KUKA KRL data list: MAIN_1.dat

&ACCESS RVP
&REL 1
&COMMENT Generated by RoboDK
&PARAM TEMPLATE = C:\KRC\Roboter\Template\vorgabe
&PARAM EDITMASK = *
DEFDAT  MAIN_1

EXT BAS (BAS_COMMAND :IN,REAL :IN )
EXT REMOTE_PROG_CALL_171()
EXT PICK_PART_111()
EXT PLACE_PART_112()
EXT EVENT_PROG_START_101()
EXT EVENT_PATH_APPROACH_102()
EXT EVENT_PATH_START_103()
EXT EVENT_PATH_FINISH_105()
EXT EVENT_PATH_RETRACT_106()
EXT EVENT_PROG_FINISH_107()
EXT PROG1_withaverylongnameandspecialcharacters()

DECL E6AXIS XP1={A1 -0.00000,A2 0.00000,A3 0.00000,A4 0.00000,A5 0.00000,A6 -0.00000}
DECL FDAT FP1={TOOL_NO 1,BASE_NO 1,IPO_FRAME #BASE,POINT2[] " ",TQ_STATE FALSE}
DECL PDAT PPDAT1={VEL 100.000,ACC 100.000,APO_DIST 1.000,APO_MODE #CPTP}
DECL E6AXIS XP2={A1 0.00000,A2 3.21124,A3 -15.42370,A4 0.00000,A5 12.21250,A6 -0.00000}
DECL FDAT FP2={TOOL_NO 1,BASE_NO 1,IPO_FRAME #BASE,POINT2[] " ",TQ_STATE FALSE}
DECL PDAT PPDAT2={VEL 100.000,ACC 100.000,APO_DIST 1.000,APO_MODE #CPTP}
DECL E6POS XP3={X 1015.000,Y 0.000,Z 1272.000,A 0.000,B 90.000,C 0.000}
DECL FDAT FP3={TOOL_NO 1,BASE_NO 1,IPO_FRAME #BASE,POINT2[] " ",TQ_STATE FALSE}
DECL LDAT LCPDAT3={VEL 1.00000,ACC 100.000,APO_DIST 1.000,APO_FAC 50.0000,ORI_TYP #VAR,CIRC_TYP #BASE,JERK_FAC 50.0000}
DECL E6AXIS XP4={A1 -29.33220,A2 46.67700,A3 -0.02452,A4 26.54560,A5 25.39570,A6 -51.63400}
DECL FDAT FP4={TOOL_NO 1,BASE_NO 1,IPO_FRAME #BASE,POINT2[] " ",TQ_STATE FALSE}
DECL PDAT PPDAT4={VEL 100.000,ACC 100.000,APO_DIST 10.000,APO_MODE #CPTP}
DECL E6POS XP5={X 187.786,Y 125.499,Z 139.112,A -179.997,B 0.180,C 179.996}
DECL FDAT FP5={TOOL_NO 1,BASE_NO 1,IPO_FRAME #BASE,POINT2[] " ",TQ_STATE FALSE}
DECL LDAT LCPDAT5={VEL 0.10000,ACC 100.000,APO_DIST 1.000,APO_FAC 50.0000,ORI_TYP #VAR,CIRC_TYP #BASE,JERK_FAC 50.0000}
DECL E6POS XP6={X 187.272,Y 447.522,Z 305.347,A 179.999,B 0.185,C -179.998}
DECL FDAT FP6={TOOL_NO 1,BASE_NO 1,IPO_FRAME #BASE,POINT2[] " ",TQ_STATE FALSE}
DECL LDAT LCPDAT6={VEL 0.30000,ACC 100.000,APO_DIST 10.000,APO_FAC 50.0000,ORI_TYP #VAR,CIRC_TYP #BASE,JERK_FAC 50.0000}
DECL E6POS XP7={X 187.851,Y 447.517,Z 126.235,A 179.999,B 0.185,C -179.998}
DECL FDAT FP7={TOOL_NO 1,BASE_NO 1,IPO_FRAME #BASE,POINT2[] " ",TQ_STATE FALSE}
DECL LDAT LCPDAT7={VEL 0.10000,ACC 100.000,APO_DIST 1.000,APO_FAC 50.0000,ORI_TYP #VAR,CIRC_TYP #BASE,JERK_FAC 50.0000}
DECL E6POS XP8={X 187.272,Y 447.522,Z 305.347,A 179.999,B 0.185,C -179.998}
DECL FDAT FP8={TOOL_NO 1,BASE_NO 1,IPO_FRAME #BASE,POINT2[] " ",TQ_STATE FALSE}
DECL LDAT LCPDAT8={VEL 0.10000,ACC 100.000,APO_DIST 10.000,APO_FAC 50.0000,ORI_TYP #VAR,CIRC_TYP #BASE,JERK_FAC 50.0000}
DECL E6AXIS XP9={A1 52.18600,A2 45.67580,A3 6.92000,A4 66.73420,A5 19.93230,A6 -92.73000}
DECL FDAT FP9={TOOL_NO 1,BASE_NO 1,IPO_FRAME #BASE,POINT2[] " ",TQ_STATE FALSE}
DECL PDAT PPDAT9={VEL 100.000,ACC 100.000,APO_DIST 25.000,APO_MODE #CPTP}
DECL E6POS XP10={X 430.047,Y 43.774,Z 231.503,A -134.549,B 11.181,C 178.913}
DECL E6POS XP11={X 109.688,Y -153.222,Z 161.073,A -134.549,B 11.181,C 178.913}
DECL FDAT FP11={TOOL_NO 1,BASE_NO 1,IPO_FRAME #BASE,POINT2[] " ",TQ_STATE FALSE}
DECL LDAT LCPDAT11={VEL 0.10000,ACC 100.000,APO_DIST 25.000,APO_FAC 50.0000,ORI_TYP #VAR,CIRC_TYP #BASE,JERK_FAC 50.0000}
DECL E6POS XP12={X 312.208,Y 292.214,Z 255.156,A -134.549,B 11.181,C 178.913}
DECL FDAT FP12={TOOL_NO 1,BASE_NO 1,IPO_FRAME #BASE,POINT2[] " ",TQ_STATE FALSE}
DECL LDAT LCPDAT12={VEL 0.10000,ACC 100.000,APO_DIST 1.000,APO_FAC 50.0000,ORI_TYP #VAR,CIRC_TYP #BASE,JERK_FAC 50.0000}
DECL E6AXIS XP13={A1 -0.00000,A2 0.00000,A3 0.00000,A4 0.00000,A5 0.00000,A6 -0.00000}
DECL FDAT FP13={TOOL_NO 1,BASE_NO 1,IPO_FRAME #BASE,POINT2[] " ",TQ_STATE FALSE}
DECL PDAT PPDAT13={VEL 100.000,ACC 100.000,APO_DIST 1.000,APO_MODE #CPTP}
DECL E6AXIS XP14={A1 88.67600,A2 29.60160,A3 -6.42883,A4 -1.98422,A5 49.47920,A6 4.54769}
DECL FDAT FP14={TOOL_NO 1,BASE_NO 1,IPO_FRAME #BASE,POINT2[] " ",TQ_STATE FALSE}
DECL PDAT PPDAT14={VEL 100.000,ACC 100.000,APO_DIST 1.000,APO_MODE #CPTP}
DECL E6POS XP15={X 19.898,Y 174.307,Z 19.008,A -94.928,B -5.426,C -179.533}
DECL FDAT FP15={TOOL_NO 1,BASE_NO 1,IPO_FRAME #BASE,POINT2[] " ",TQ_STATE FALSE}
DECL LDAT LCPDAT15={VEL 0.10000,ACC 100.000,APO_DIST 1.000,APO_FAC 50.0000,ORI_TYP #VAR,CIRC_TYP #BASE,JERK_FAC 50.0000}
DECL E6POS XP16={X 378.402,Y 174.416,Z 18.997,A -94.928,B -5.426,C -179.533}
DECL FDAT FP16={TOOL_NO 1,BASE_NO 1,IPO_FRAME #BASE,POINT2[] " ",TQ_STATE FALSE}
DECL LDAT LCPDAT16={VEL 0.10000,ACC 100.000,APO_DIST 1.000,APO_FAC 50.0000,ORI_TYP #VAR,CIRC_TYP #BASE,JERK_FAC 50.0000}
DECL E6POS XP17={X 380.996,Y 112.363,Z 34.882,A -95.294,B -18.136,C -178.348}
DECL FDAT FP17={TOOL_NO 1,BASE_NO 1,IPO_FRAME #BASE,POINT2[] " ",TQ_STATE FALSE}
DECL LDAT LCPDAT17={VEL 0.10000,ACC 100.000,APO_DIST 1.000,APO_FAC 50.0000,ORI_TYP #VAR,CIRC_TYP #BASE,JERK_FAC 50.0000}
DECL E6POS XP18={X 16.551,Y 114.359,Z 34.226,A -95.294,B -18.136,C -178.348}
DECL FDAT FP18={TOOL_NO 1,BASE_NO 1,IPO_FRAME #BASE,POINT2[] " ",TQ_STATE FALSE}
DECL LDAT LCPDAT18={VEL 0.10000,ACC 100.000,APO_DIST 1.000,APO_FAC 50.0000,ORI_TYP #VAR,CIRC_TYP #BASE,JERK_FAC 50.0000}
DECL E6POS XP19={X 26.434,Y 54.524,Z 46.072,A -95.461,B 4.348,C 179.585}
DECL FDAT FP19={TOOL_NO 1,BASE_NO 1,IPO_FRAME #BASE,POINT2[] " ",TQ_STATE FALSE}
DECL LDAT LCPDAT19={VEL 0.10000,ACC 100.000,APO_DIST 1.000,APO_FAC 50.0000,ORI_TYP #VAR,CIRC_TYP #BASE,JERK_FAC 50.0000}
DECL E6POS XP20={X 385.448,Y 48.050,Z 45.137,A -95.590,B 11.181,C 178.913}
DECL FDAT FP20={TOOL_NO 1,BASE_NO 1,IPO_FRAME #BASE,POINT2[] " ",TQ_STATE FALSE}
DECL LDAT LCPDAT20={VEL 0.10000,ACC 100.000,APO_DIST 1.000,APO_FAC 50.0000,ORI_TYP #VAR,CIRC_TYP #BASE,JERK_FAC 50.0000}
DECL E6POS XP21={X 385.448,Y -1.625,Z 295.251,A -95.590,B 11.181,C 178.913}
DECL FDAT FP21={TOOL_NO 1,BASE_NO 1,IPO_FRAME #BASE,POINT2[] " ",TQ_STATE FALSE}
DECL LDAT LCPDAT21={VEL 0.10000,ACC 100.000,APO_DIST 1.000,APO_FAC 50.0000,ORI_TYP #VAR,CIRC_TYP #BASE,JERK_FAC 50.0000}
DECL E6AXIS XP22={A1 -0.00000,A2 0.00000,A3 0.00000,A4 0.00000,A5 0.00000,A6 -0.00000}
DECL FDAT FP22={TOOL_NO 1,BASE_NO 1,IPO_FRAME #BASE,POINT2[] " ",TQ_STATE FALSE}
DECL PDAT PPDAT22={VEL 100.000,ACC 100.000,APO_DIST 1.000,APO_MODE #CPTP}
DECL E6AXIS XP23={A1 -68.09030,A2 24.20190,A3 26.78550,A4 38.21340,A5 36.20170,A6 -98.79640}
DECL FDAT FP23={TOOL_NO 1,BASE_NO 1,IPO_FRAME #BASE,POINT2[] " ",TQ_STATE FALSE}
DECL PDAT PPDAT23={VEL 100.000,ACC 100.000,APO_DIST 1.000,APO_MODE #CPTP}
DECL E6POS XP24={X -49.895,Y 253.259,Z 319.999,A -90.000,B 0.353,C -179.975}
DECL FDAT FP24={TOOL_NO 1,BASE_NO 1,IPO_FRAME #BASE,POINT2[] " ",TQ_STATE FALSE}
DECL LDAT LCPDAT24={VEL 1.00000,ACC 100.000,APO_DIST 1.000,APO_FAC 50.0000,ORI_TYP #VAR,CIRC_TYP #BASE,JERK_FAC 50.0000}
DECL E6POS XP25={X 0.000,Y 250.000,Z 270.000,A -90.000,B 0.353,C -179.975}
DECL FDAT FP25={TOOL_NO 1,BASE_NO 1,IPO_FRAME #BASE,POINT2[] " ",TQ_STATE FALSE}
DECL LDAT LCPDAT25={VEL 1.00000,ACC 100.000,APO_DIST 1.000,APO_FAC 50.0000,ORI_TYP #VAR,CIRC_TYP #BASE,JERK_FAC 50.0000}
DECL E6POS XP26={X 35.579,Y 247.455,Z 270.000,A -90.000,B 0.345,C -179.925}
DECL FDAT FP26={TOOL_NO 1,BASE_NO 1,IPO_FRAME #BASE,POINT2[] " ",TQ_STATE FALSE}
DECL LDAT LCPDAT26={VEL 0.05000,ACC 100.000,APO_DIST 1.000,APO_FAC 50.0000,ORI_TYP #VAR,CIRC_TYP #BASE,JERK_FAC 50.0000}
DECL E6POS XP27={X 70.433,Y 239.873,Z 270.000,A -89.999,B 0.331,C -179.876}
DECL FDAT FP27={TOOL_NO 1,BASE_NO 1,IPO_FRAME #BASE,POINT2[] " ",TQ_STATE FALSE}
DECL LDAT LCPDAT27={VEL 0.05000,ACC 100.000,APO_DIST 1.000,APO_FAC 50.0000,ORI_TYP #VAR,CIRC_TYP #BASE,JERK_FAC 50.0000}
DECL E6POS XP28={X 103.854,Y 227.408,Z 270.000,A -89.999,B 0.310,C -179.831}
DECL FDAT FP28={TOOL_NO 1,BASE_NO 1,IPO_FRAME #BASE,POINT2[] " ",TQ_STATE FALSE}
DECL LDAT LCPDAT28={VEL 0.05000,ACC 100.000,APO_DIST 1.000,APO_FAC 50.0000,ORI_TYP #VAR,CIRC_TYP #BASE,JERK_FAC 50.0000}
DECL E6POS XP29={X 135.160,Y 210.313,Z 270.000,A -89.999,B 0.283,C -179.788}
DECL FDAT FP29={TOOL_NO 1,BASE_NO 1,IPO_FRAME #BASE,POINT2[] " ",TQ_STATE FALSE}
DECL LDAT LCPDAT29={VEL 0.05000,ACC 100.000,APO_DIST 1.000,APO_FAC 50.0000,ORI_TYP #VAR,CIRC_TYP #BASE,JERK_FAC 50.0000}
DECL E6POS XP30={X 163.715,Y 188.937,Z 270.000,A -89.999,B 0.250,C -179.750}
DECL FDAT FP30={TOOL_NO 1,BASE_NO 1,IPO_FRAME #BASE,POINT2[] " ",TQ_STATE FALSE}
DECL LDAT LCPDAT30={VEL 0.05000,ACC 100.000,APO_DIST 1.000,APO_FAC 50.0000,ORI_TYP #VAR,CIRC_TYP #BASE,JERK_FAC 50.0000}
DECL E6POS XP31={X 188.937,Y 163.715,Z 270.000,A -89.999,B 0.212,C -179.717}
DECL FDAT FP31={TOOL_NO 1,BASE_NO 1,IPO_FRAME #BASE,POINT2[] " ",TQ_STATE FALSE}
DECL LDAT LCPDAT31={VEL 0.05000,ACC 100.000,APO_DIST 1.000,APO_FAC 50.0000,ORI_TYP #VAR,CIRC_TYP #BASE,JERK_FAC 50.0000}
DECL E6POS XP32={X 210.313,Y 135.160,Z 270.000,A -89.999,B 0.170,C -179.689}
DECL FDAT FP32={TOOL_NO 1,BASE_NO 1,IPO_FRAME #BASE,POINT2[] " ",TQ_STATE FALSE}
DECL LDAT LCPDAT32={VEL 0.05000,ACC 100.000,APO_DIST 1.000,APO_FAC 50.0000,ORI_TYP #VAR,CIRC_TYP #BASE,JERK_FAC 50.0000}
DECL E6POS XP33={X 227.408,Y 103.854,Z 270.000,A -89.999,B 0.124,C -179.668}
DECL FDAT FP33={TOOL_NO 1,BASE_NO 1,IPO_FRAME #BASE,POINT2[] " ",TQ_STATE FALSE}
DECL LDAT LCPDAT33={VEL 0.05000,ACC 100.000,APO_DIST 1.000,APO_FAC 50.0000,ORI_TYP #VAR,CIRC_TYP #BASE,JERK_FAC 50.0000}
DECL E6POS XP34={X 239.873,Y 70.433,Z 270.000,A -90.000,B 0.075,C -179.654}
DECL FDAT FP34={TOOL_NO 1,BASE_NO 1,IPO_FRAME #BASE,POINT2[] " ",TQ_STATE FALSE}
DECL LDAT LCPDAT34={VEL 0.05000,ACC 100.000,APO_DIST 1.000,APO_FAC 50.0000,ORI_TYP #VAR,CIRC_TYP #BASE,JERK_FAC 50.0000}
DECL E6POS XP35={X 247.455,Y 35.579,Z 270.000,A -90.000,B 0.025,C -179.647}
DECL FDAT FP35={TOOL_NO 1,BASE_NO 1,IPO_FRAME #BASE,POINT2[] " ",TQ_STATE FALSE}
DECL LDAT LCPDAT35={VEL 0.05000,ACC 100.000,APO_DIST 1.000,APO_FAC 50.0000,ORI_TYP #VAR,CIRC_TYP #BASE,JERK_FAC 50.0000}
DECL E6POS XP36={X 250.000,Y 0.000,Z 270.000,A -90.000,B -0.025,C -179.647}
DECL FDAT FP36={TOOL_NO 1,BASE_NO 1,IPO_FRAME #BASE,POINT2[] " ",TQ_STATE FALSE}
DECL LDAT LCPDAT36={VEL 0.05000,ACC 100.000,APO_DIST 1.000,APO_FAC 50.0000,ORI_TYP #VAR,CIRC_TYP #BASE,JERK_FAC 50.0000}
DECL E6POS XP37={X 247.455,Y -35.579,Z 270.000,A -90.000,B -0.075,C -179.654}
DECL FDAT FP37={TOOL_NO 1,BASE_NO 1,IPO_FRAME #BASE,POINT2[] " ",TQ_STATE FALSE}
DECL LDAT LCPDAT37={VEL 0.05000,ACC 100.000,APO_DIST 1.000,APO_FAC 50.0000,ORI_TYP #VAR,CIRC_TYP #BASE,JERK_FAC 50.0000}
DECL E6POS XP38={X 239.873,Y -70.433,Z 270.000,A -90.001,B -0.124,C -179.668}
DECL FDAT FP38={TOOL_NO 1,BASE_NO 1,IPO_FRAME #BASE,POINT2[] " ",TQ_STATE FALSE}
DECL LDAT LCPDAT38={VEL 0.05000,ACC 100.000,APO_DIST 1.000,APO_FAC 50.0000,ORI_TYP #VAR,CIRC_TYP #BASE,JERK_FAC 50.0000}
DECL E6POS XP39={X 227.408,Y -103.854,Z 270.000,A -90.001,B -0.170,C -179.689}
DECL FDAT FP39={TOOL_NO 1,BASE_NO 1,IPO_FRAME #BASE,POINT2[] " ",TQ_STATE FALSE}
DECL LDAT LCPDAT39={VEL 0.05000,ACC 100.000,APO_DIST 1.000,APO_FAC 50.0000,ORI_TYP #VAR,CIRC_TYP #BASE,JERK_FAC 50.0000}
DECL E6POS XP40={X 210.313,Y -135.160,Z 270.000,A -90.001,B -0.212,C -179.717}
DECL FDAT FP40={TOOL_NO 1,BASE_NO 1,IPO_FRAME #BASE,POINT2[] " ",TQ_STATE FALSE}
DECL LDAT LCPDAT40={VEL 0.05000,ACC 100.000,APO_DIST 1.000,APO_FAC 50.0000,ORI_TYP #VAR,CIRC_TYP #BASE,JERK_FAC 50.0000}
DECL E6POS XP41={X 188.937,Y -163.715,Z 270.000,A -90.001,B -0.250,C -179.750}
DECL FDAT FP41={TOOL_NO 1,BASE_NO 1,IPO_FRAME #BASE,POINT2[] " ",TQ_STATE FALSE}
DECL LDAT LCPDAT41={VEL 0.05000,ACC 100.000,APO_DIST 1.000,APO_FAC 50.0000,ORI_TYP #VAR,CIRC_TYP #BASE,JERK_FAC 50.0000}
DECL E6POS XP42={X 163.715,Y -188.937,Z 270.000,A -90.001,B -0.283,C -179.788}
DECL FDAT FP42={TOOL_NO 1,BASE_NO 1,IPO_FRAME #BASE,POINT2[] " ",TQ_STATE FALSE}
DECL LDAT LCPDAT42={VEL 0.05000,ACC 100.000,APO_DIST 1.000,APO_FAC 50.0000,ORI_TYP #VAR,CIRC_TYP #BASE,JERK_FAC 50.0000}
DECL E6POS XP43={X 135.160,Y -210.313,Z 270.000,A -90.001,B -0.311,C -179.830}
DECL FDAT FP43={TOOL_NO 1,BASE_NO 1,IPO_FRAME #BASE,POINT2[] " ",TQ_STATE FALSE}
DECL LDAT LCPDAT43={VEL 0.05000,ACC 100.000,APO_DIST 1.000,APO_FAC 50.0000,ORI_TYP #VAR,CIRC_TYP #BASE,JERK_FAC 50.0000}
DECL E6POS XP44={X 103.854,Y -227.408,Z 270.000,A -90.001,B -0.332,C -179.876}
DECL FDAT FP44={TOOL_NO 1,BASE_NO 1,IPO_FRAME #BASE,POINT2[] " ",TQ_STATE FALSE}
DECL LDAT LCPDAT44={VEL 0.05000,ACC 100.000,APO_DIST 1.000,APO_FAC 50.0000,ORI_TYP #VAR,CIRC_TYP #BASE,JERK_FAC 50.0000}
DECL E6POS XP45={X 70.433,Y -239.873,Z 270.000,A -90.000,B -0.346,C -179.925}
DECL FDAT FP45={TOOL_NO 1,BASE_NO 1,IPO_FRAME #BASE,POINT2[] " ",TQ_STATE FALSE}
DECL LDAT LCPDAT45={VEL 0.05000,ACC 100.000,APO_DIST 1.000,APO_FAC 50.0000,ORI_TYP #VAR,CIRC_TYP #BASE,JERK_FAC 50.0000}
DECL E6POS XP46={X 35.579,Y -247.455,Z 270.000,A -90.000,B -0.353,C -179.975}
DECL FDAT FP46={TOOL_NO 1,BASE_NO 1,IPO_FRAME #BASE,POINT2[] " ",TQ_STATE FALSE}
DECL LDAT LCPDAT46={VEL 0.05000,ACC 100.000,APO_DIST 1.000,APO_FAC 50.0000,ORI_TYP #VAR,CIRC_TYP #BASE,JERK_FAC 50.0000}
DECL E6POS XP47={X 0.000,Y -250.000,Z 270.000,A -90.000,B -0.353,C -179.975}
DECL FDAT FP47={TOOL_NO 1,BASE_NO 1,IPO_FRAME #BASE,POINT2[] " ",TQ_STATE FALSE}
DECL LDAT LCPDAT47={VEL 0.05000,ACC 100.000,APO_DIST 1.000,APO_FAC 50.0000,ORI_TYP #VAR,CIRC_TYP #BASE,JERK_FAC 50.0000}
DECL E6POS XP48={X 0.000,Y -250.000,Z 270.000,A -90.000,B -0.353,C 179.975}
DECL FDAT FP48={TOOL_NO 1,BASE_NO 1,IPO_FRAME #BASE,POINT2[] " ",TQ_STATE FALSE}
DECL LDAT LCPDAT48={VEL 0.05000,ACC 100.000,APO_DIST 1.000,APO_FAC 50.0000,ORI_TYP #VAR,CIRC_TYP #BASE,JERK_FAC 50.0000}
DECL E6POS XP49={X -35.579,Y -247.455,Z 270.000,A -90.000,B -0.346,C 179.925}
DECL FDAT FP49={TOOL_NO 1,BASE_NO 1,IPO_FRAME #BASE,POINT2[] " ",TQ_STATE FALSE}
DECL LDAT LCPDAT49={VEL 0.05000,ACC 100.000,APO_DIST 1.000,APO_FAC 50.0000,ORI_TYP #VAR,CIRC_TYP #BASE,JERK_FAC 50.0000}
DECL E6POS XP50={X -70.433,Y -239.873,Z 270.000,A -89.999,B -0.331,C 179.876}
DECL FDAT FP50={TOOL_NO 1,BASE_NO 1,IPO_FRAME #BASE,POINT2[] " ",TQ_STATE FALSE}
DECL LDAT LCPDAT50={VEL 0.05000,ACC 100.000,APO_DIST 1.000,APO_FAC 50.0000,ORI_TYP #VAR,CIRC_TYP #BASE,JERK_FAC 50.0000}
DECL E6POS XP51={X -103.854,Y -227.408,Z 270.000,A -89.999,B -0.310,C 179.831}
DECL FDAT FP51={TOOL_NO 1,BASE_NO 1,IPO_FRAME #BASE,POINT2[] " ",TQ_STATE FALSE}
DECL LDAT LCPDAT51={VEL 0.05000,ACC 100.000,APO_DIST 1.000,APO_FAC 50.0000,ORI_TYP #VAR,CIRC_TYP #BASE,JERK_FAC 50.0000}
DECL E6POS XP52={X -135.160,Y -210.313,Z 270.000,A -89.999,B -0.283,C 179.788}
DECL FDAT FP52={TOOL_NO 1,BASE_NO 1,IPO_FRAME #BASE,POINT2[] " ",TQ_STATE FALSE}
DECL LDAT LCPDAT52={VEL 0.05000,ACC 100.000,APO_DIST 1.000,APO_FAC 50.0000,ORI_TYP #VAR,CIRC_TYP #BASE,JERK_FAC 50.0000}
DECL E6POS XP53={X -163.715,Y -188.937,Z 270.000,A -89.999,B -0.250,C 179.750}
DECL FDAT FP53={TOOL_NO 1,BASE_NO 1,IPO_FRAME #BASE,POINT2[] " ",TQ_STATE FALSE}
DECL LDAT LCPDAT53={VEL 0.05000,ACC 100.000,APO_DIST 1.000,APO_FAC 50.0000,ORI_TYP #VAR,CIRC_TYP #BASE,JERK_FAC 50.0000}
DECL E6POS XP54={X -188.937,Y -163.715,Z 270.000,A -89.999,B -0.212,C 179.717}
DECL FDAT FP54={TOOL_NO 1,BASE_NO 1,IPO_FRAME #BASE,POINT2[] " ",TQ_STATE FALSE}
DECL LDAT LCPDAT54={VEL 0.05000,ACC 100.000,APO_DIST 1.000,APO_FAC 50.0000,ORI_TYP #VAR,CIRC_TYP #BASE,JERK_FAC 50.0000}
DECL E6POS XP55={X -210.313,Y -135.160,Z 270.000,A -89.999,B -0.169,C 179.690}
DECL FDAT FP55={TOOL_NO 1,BASE_NO 1,IPO_FRAME #BASE,POINT2[] " ",TQ_STATE FALSE}
DECL LDAT LCPDAT55={VEL 0.05000,ACC 100.000,APO_DIST 1.000,APO_FAC 50.0000,ORI_TYP #VAR,CIRC_TYP #BASE,JERK_FAC 50.0000}
DECL E6POS XP56={X -227.408,Y -103.854,Z 270.000,A -89.999,B -0.123,C 179.669}
DECL FDAT FP56={TOOL_NO 1,BASE_NO 1,IPO_FRAME #BASE,POINT2[] " ",TQ_STATE FALSE}
DECL LDAT LCPDAT56={VEL 0.05000,ACC 100.000,APO_DIST 1.000,APO_FAC 50.0000,ORI_TYP #VAR,CIRC_TYP #BASE,JERK_FAC 50.0000}
DECL E6POS XP57={X -239.873,Y -70.433,Z 270.000,A -90.000,B -0.075,C 179.654}
DECL FDAT FP57={TOOL_NO 1,BASE_NO 1,IPO_FRAME #BASE,POINT2[] " ",TQ_STATE FALSE}
DECL LDAT LCPDAT57={VEL 0.05000,ACC 100.000,APO_DIST 1.000,APO_FAC 50.0000,ORI_TYP #VAR,CIRC_TYP #BASE,JERK_FAC 50.0000}
DECL E6POS XP58={X -247.455,Y -35.579,Z 270.000,A -90.000,B -0.025,C 179.647}
DECL FDAT FP58={TOOL_NO 1,BASE_NO 1,IPO_FRAME #BASE,POINT2[] " ",TQ_STATE FALSE}
DECL LDAT LCPDAT58={VEL 0.05000,ACC 100.000,APO_DIST 1.000,APO_FAC 50.0000,ORI_TYP #VAR,CIRC_TYP #BASE,JERK_FAC 50.0000}
DECL E6POS XP59={X -250.000,Y 0.000,Z 270.000,A -90.000,B 0.025,C 179.647}
DECL FDAT FP59={TOOL_NO 1,BASE_NO 1,IPO_FRAME #BASE,POINT2[] " ",TQ_STATE FALSE}
DECL LDAT LCPDAT59={VEL 0.05000,ACC 100.000,APO_DIST 1.000,APO_FAC 50.0000,ORI_TYP #VAR,CIRC_TYP #BASE,JERK_FAC 50.0000}
DECL E6POS XP60={X -247.455,Y 35.579,Z 270.000,A -90.000,B 0.075,C 179.655}
DECL FDAT FP60={TOOL_NO 1,BASE_NO 1,IPO_FRAME #BASE,POINT2[] " ",TQ_STATE FALSE}
DECL LDAT LCPDAT60={VEL 0.05000,ACC 100.000,APO_DIST 1.000,APO_FAC 50.0000,ORI_TYP #VAR,CIRC_TYP #BASE,JERK_FAC 50.0000}
DECL E6POS XP61={X -239.873,Y 70.433,Z 270.000,A -90.001,B 0.123,C 179.669}
DECL FDAT FP61={TOOL_NO 1,BASE_NO 1,IPO_FRAME #BASE,POINT2[] " ",TQ_STATE FALSE}
DECL LDAT LCPDAT61={VEL 0.05000,ACC 100.000,APO_DIST 1.000,APO_FAC 50.0000,ORI_TYP #VAR,CIRC_TYP #BASE,JERK_FAC 50.0000}
DECL E6POS XP62={X -227.408,Y 103.854,Z 270.000,A -90.001,B 0.170,C 179.689}
DECL FDAT FP62={TOOL_NO 1,BASE_NO 1,IPO_FRAME #BASE,POINT2[] " ",TQ_STATE FALSE}
DECL LDAT LCPDAT62={VEL 0.05000,ACC 100.000,APO_DIST 1.000,APO_FAC 50.0000,ORI_TYP #VAR,CIRC_TYP #BASE,JERK_FAC 50.0000}
DECL E6POS XP63={X -210.313,Y 135.160,Z 270.000,A -90.001,B 0.212,C 179.717}
DECL FDAT FP63={TOOL_NO 1,BASE_NO 1,IPO_FRAME #BASE,POINT2[] " ",TQ_STATE FALSE}
DECL LDAT LCPDAT63={VEL 0.05000,ACC 100.000,APO_DIST 1.000,APO_FAC 50.0000,ORI_TYP #VAR,CIRC_TYP #BASE,JERK_FAC 50.0000}
DECL E6POS XP64={X -188.937,Y 163.715,Z 270.000,A -90.001,B 0.250,C 179.750}
DECL FDAT FP64={TOOL_NO 1,BASE_NO 1,IPO_FRAME #BASE,POINT2[] " ",TQ_STATE FALSE}
DECL LDAT LCPDAT64={VEL 0.05000,ACC 100.000,APO_DIST 1.000,APO_FAC 50.0000,ORI_TYP #VAR,CIRC_TYP #BASE,JERK_FAC 50.0000}
DECL E6POS XP65={X -163.715,Y 188.937,Z 270.000,A -90.001,B 0.283,C 179.788}
DECL FDAT FP65={TOOL_NO 1,BASE_NO 1,IPO_FRAME #BASE,POINT2[] " ",TQ_STATE FALSE}
DECL LDAT LCPDAT65={VEL 0.05000,ACC 100.000,APO_DIST 1.000,APO_FAC 50.0000,ORI_TYP #VAR,CIRC_TYP #BASE,JERK_FAC 50.0000}
DECL E6POS XP66={X -135.160,Y 210.313,Z 270.000,A -90.001,B 0.310,C 179.831}
DECL FDAT FP66={TOOL_NO 1,BASE_NO 1,IPO_FRAME #BASE,POINT2[] " ",TQ_STATE FALSE}
DECL LDAT LCPDAT66={VEL 0.05000,ACC 100.000,APO_DIST 1.000,APO_FAC 50.0000,ORI_TYP #VAR,CIRC_TYP #BASE,JERK_FAC 50.0000}
DECL E6POS XP67={X -103.854,Y 227.408,Z 270.000,A -90.001,B 0.332,C 179.876}
DECL FDAT FP67={TOOL_NO 1,BASE_NO 1,IPO_FRAME #BASE,POINT2[] " ",TQ_STATE FALSE}
DECL LDAT LCPDAT67={VEL 0.05000,ACC 100.000,APO_DIST 1.000,APO_FAC 50.0000,ORI_TYP #VAR,CIRC_TYP #BASE,JERK_FAC 50.0000}
DECL E6POS XP68={X -70.433,Y 239.873,Z 270.000,A -90.000,B 0.346,C 179.925}
DECL FDAT FP68={TOOL_NO 1,BASE_NO 1,IPO_FRAME #BASE,POINT2[] " ",TQ_STATE FALSE}
DECL LDAT LCPDAT68={VEL 0.05000,ACC 100.000,APO_DIST 1.000,APO_FAC 50.0000,ORI_TYP #VAR,CIRC_TYP #BASE,JERK_FAC 50.0000}
DECL E6POS XP69={X -35.579,Y 247.455,Z 270.000,A -90.000,B 0.353,C 179.975}
DECL FDAT FP69={TOOL_NO 1,BASE_NO 1,IPO_FRAME #BASE,POINT2[] " ",TQ_STATE FALSE}
DECL LDAT LCPDAT69={VEL 0.05000,ACC 100.000,APO_DIST 1.000,APO_FAC 50.0000,ORI_TYP #VAR,CIRC_TYP #BASE,JERK_FAC 50.0000}
DECL E6POS XP70={X 0.000,Y 250.000,Z 270.000,A -90.000,B 0.353,C 179.975}
DECL FDAT FP70={TOOL_NO 1,BASE_NO 1,IPO_FRAME #BASE,POINT2[] " ",TQ_STATE FALSE}
DECL LDAT LCPDAT70={VEL 0.05000,ACC 100.000,APO_DIST 1.000,APO_FAC 50.0000,ORI_TYP #VAR,CIRC_TYP #BASE,JERK_FAC 50.0000}
DECL E6POS XP71={X 49.895,Y 253.258,Z 319.999,A -90.000,B 0.353,C 179.975}
DECL FDAT FP71={TOOL_NO 1,BASE_NO 1,IPO_FRAME #BASE,POINT2[] " ",TQ_STATE FALSE}
DECL LDAT LCPDAT71={VEL 1.00000,ACC 100.000,APO_DIST 1.000,APO_FAC 50.0000,ORI_TYP #VAR,CIRC_TYP #BASE,JERK_FAC 50.0000}
DECL E6POS XP72={X 49.939,Y 252.642,Z 419.997,A -90.000,B 0.353,C 179.975}
DECL FDAT FP72={TOOL_NO 1,BASE_NO 1,IPO_FRAME #BASE,POINT2[] " ",TQ_STATE FALSE}
DECL LDAT LCPDAT72={VEL 1.00000,ACC 100.000,APO_DIST 1.000,APO_FAC 50.0000,ORI_TYP #VAR,CIRC_TYP #BASE,JERK_FAC 50.0000}
DECL E6AXIS XP73={A1 -29.33220,A2 46.67700,A3 -0.02452,A4 26.54560,A5 25.39570,A6 -51.63400}
DECL FDAT FP73={TOOL_NO 1,BASE_NO 1,IPO_FRAME #BASE,POINT2[] " ",TQ_STATE FALSE}
DECL PDAT PPDAT73={VEL 100.000,ACC 100.000,APO_DIST 1.000,APO_MODE #CPTP}
DECL E6POS XP74={X 187.786,Y 125.499,Z 139.112,A -179.997,B 0.180,C 179.996}
DECL FDAT FP74={TOOL_NO 1,BASE_NO 1,IPO_FRAME #BASE,POINT2[] " ",TQ_STATE FALSE}
DECL LDAT LCPDAT74={VEL 1.00000,ACC 100.000,APO_DIST 1.000,APO_FAC 50.0000,ORI_TYP #VAR,CIRC_TYP #BASE,JERK_FAC 50.0000}
DECL E6POS XP75={X 187.264,Y 125.487,Z 305.356,A 180.000,B 0.184,C -180.000}
DECL FDAT FP75={TOOL_NO 1,BASE_NO 1,IPO_FRAME #BASE,POINT2[] " ",TQ_STATE FALSE}
DECL LDAT LCPDAT75={VEL 1.00000,ACC 100.000,APO_DIST 1.000,APO_FAC 50.0000,ORI_TYP #VAR,CIRC_TYP #BASE,JERK_FAC 50.0000}
DECL E6AXIS XP76={A1 -0.00000,A2 0.00000,A3 0.00000,A4 0.00000,A5 0.00000,A6 -0.00000}
DECL FDAT FP76={TOOL_NO 1,BASE_NO 1,IPO_FRAME #BASE,POINT2[] " ",TQ_STATE FALSE}
DECL PDAT PPDAT76={VEL 100.000,ACC 100.000,APO_DIST 1.000,APO_MODE #CPTP}

ENDDAT
